FUNCTION_BLOCK HI_THRESHOLD
  {SET_ATTRIBUTE(OpcUa, SERVICE)}
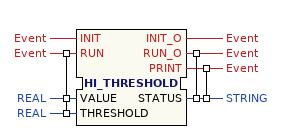
  EVENT_INPUT
    INIT;
    RUN WITH VALUE, THRESHOLD;
  END_EVENT
  EVENT_OUTPUT
    INIT_O;
    RUN_O WITH STATUS;
    PRINT WITH STATUS;
  END_EVENT
  VAR_INPUT
    VALUE : REAL; {SET_ATTRIBUTE(OpcUa, Variable)}
    THRESHOLD : REAL; {SET_ATTRIBUTE(OpcUa, Variable)}
  END_VAR
  VAR_OUTPUT
    STATUS : STRING; {SET_ATTRIBUTE(OpcUa, Variable)}
  END_VAR
END_FUNCTION_BLOCK
